Fanuc KAREL source: kc00052.KL

-- PROVISIONAL review KL for V940-1; original PC SHA256 cceacf85e9ac910581f4afd31474bd34dd836ef02914e90f7287c13185ba2a7b
-- Incomplete behavior may be omitted. Consult companion uncertainty JSON. Do not deploy.
PROGRAM KC00052
%NOLOCKGROUP
BEGIN
  -- V9_ZERO_TABLE_METADATA_HINT layout=0002_ascii; no indexed target words; source/name/runtime held
  -- UNRESOLVED_PC offsets 5-39; opcodes 27,22,22,22,22,22,31
  -- UNRESOLVED_PC offsets 44-48; opcodes 7F
END KC00052
